// Mitsubishi GX Works2 project: B_v6_v2   PLC: Q03UDE

PROGRAM COMMON
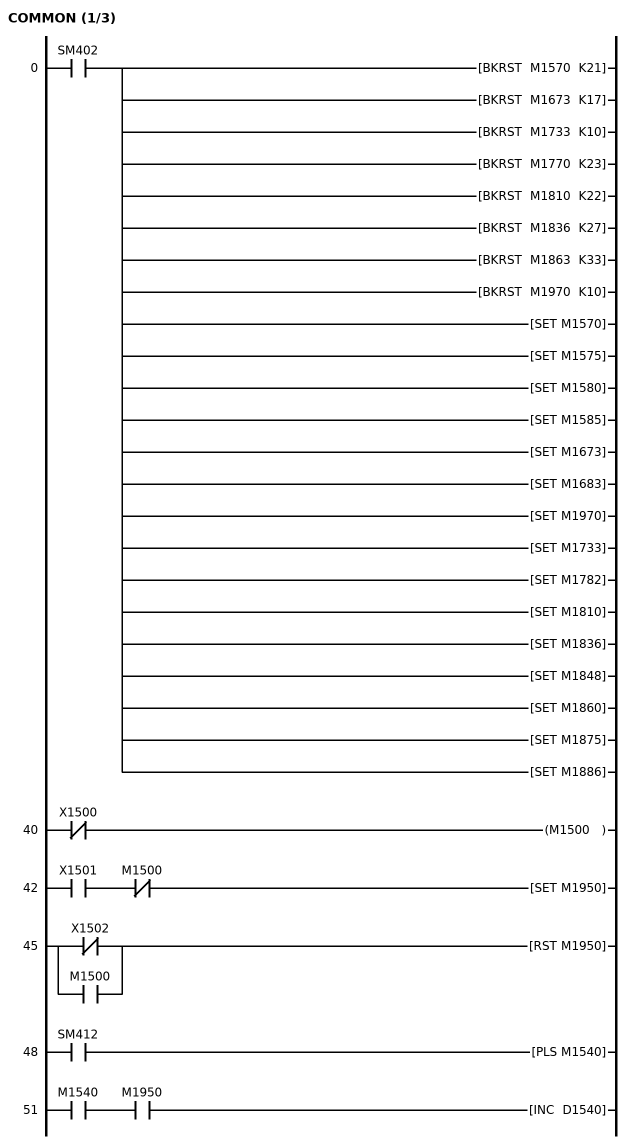
0     LD      SM402
      BKRST   M1570 K21
      BKRST   M1673 K17
      BKRST   M1733 K10
      BKRST   M1770 K23
      BKRST   M1810 K22
      BKRST   M1836 K27
      BKRST   M1863 K33
      BKRST   M1970 K10
      SET     M1570
      SET     M1575
      SET     M1580
      SET     M1585
      SET     M1673
      SET     M1683
      SET     M1970
      SET     M1733
      SET     M1782
      SET     M1810
      SET     M1836
      SET     M1848
      SET     M1860
      SET     M1875
      SET     M1886
40    LDI     X1500
      OUT     M1500
42    LD      X1501
      ANI     M1500
      SET     M1950
45    LDI     X1502
      OR      M1500
      RST     M1950
48    LD      SM412
      PLS     M1540
51    LD      M1540
      AND     M1950
      INC     D1540
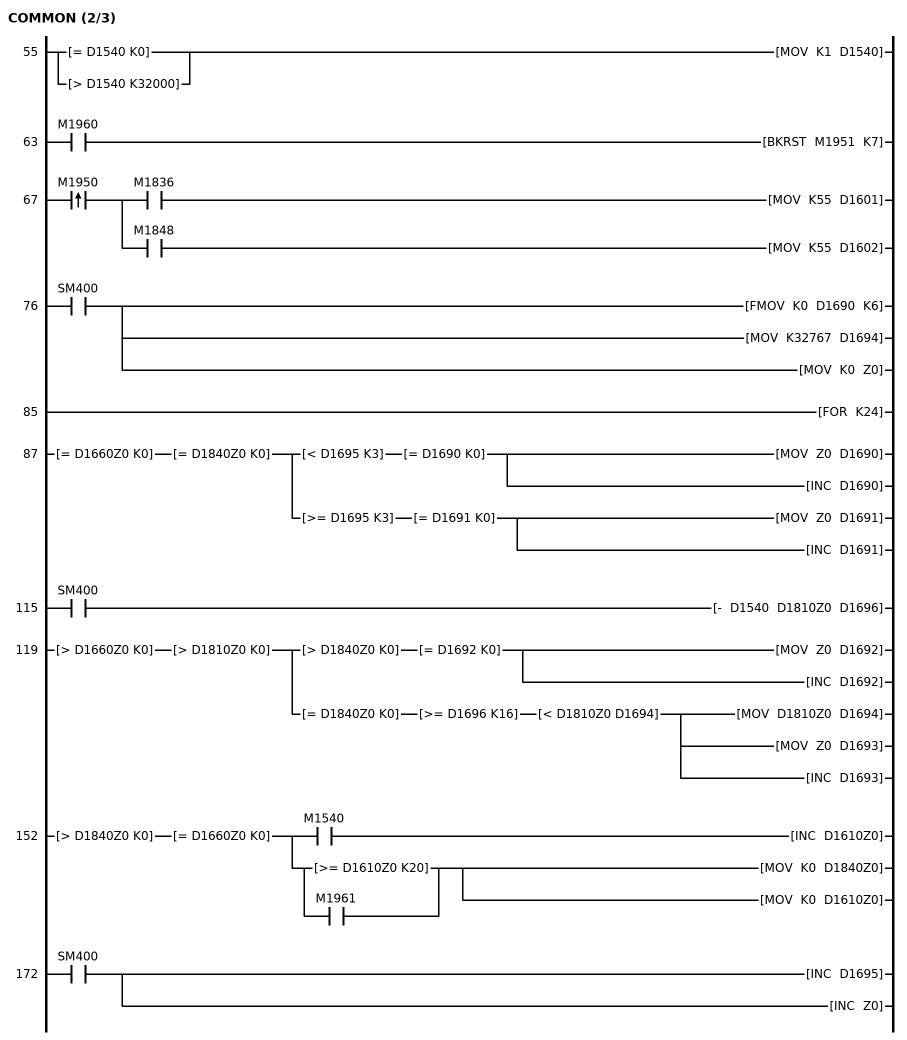
55    LD=     D1540 K0
      OR>     D1540 K32000
      MOV     K1 D1540
63    LD      M1960
      BKRST   M1951 K7
67    LDP     M1950
      MPS
      AND     M1836
      MOV     K55 D1601
      MPP
      AND     M1848
      MOV     K55 D1602
76    LD      SM400
      FMOV    K0 D1690 K6
      MOV     K32767 D1694
      MOV     K0 Z0
85    FOR     K24
87    LD=     D1660Z0 K0
      AND=    D1840Z0 K0
      MPS
      AND<    D1695 K3
      AND=    D1690 K0
      MOV     Z0 D1690
      INC     D1690
      MPP
      AND>=   D1695 K3
      AND=    D1691 K0
      MOV     Z0 D1691
      INC     D1691
115   LD      SM400
      -       D1540 D1810Z0 D1696
119   LD>     D1660Z0 K0
      AND>    D1810Z0 K0
      MPS
      AND>    D1840Z0 K0
      AND=    D1692 K0
      MOV     Z0 D1692
      INC     D1692
      MPP
      AND=    D1840Z0 K0
      AND>=   D1696 K16
      AND<    D1810Z0 D1694
      MOV     D1810Z0 D1694
      MOV     Z0 D1693
      INC     D1693
152   LD>     D1840Z0 K0
      AND=    D1660Z0 K0
      MPS
      AND     M1540
      INC     D1610Z0
      MPP
      LD>=    D1610Z0 K20
      OR      M1961
      ANB
      MOV     K0 D1840Z0
      MOV     K0 D1610Z0
172   LD      SM400
      INC     D1695
      INC     Z0
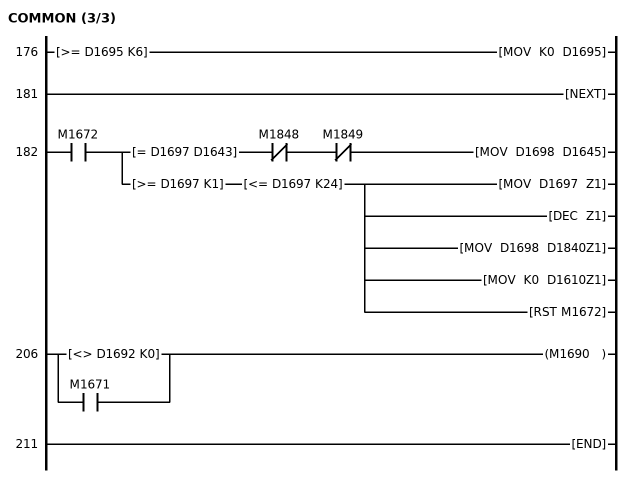
176   LD>=    D1695 K6
      MOV     K0 D1695
181   NEXT
182   LD      M1672
      MPS
      AND=    D1697 D1643
      ANI     M1848
      ANI     M1849
      MOV     D1698 D1645
      MPP
      AND>=   D1697 K1
      AND<=   D1697 K24
      MOV     D1697 Z1
      DEC     Z1
      MOV     D1698 D1840Z1
      MOV     K0 D1610Z1
      RST     M1672
206   LD<>    D1692 K0
      OR      M1671
      OUT     M1690
211   END
END_PROGRAM

PROGRAM RFID
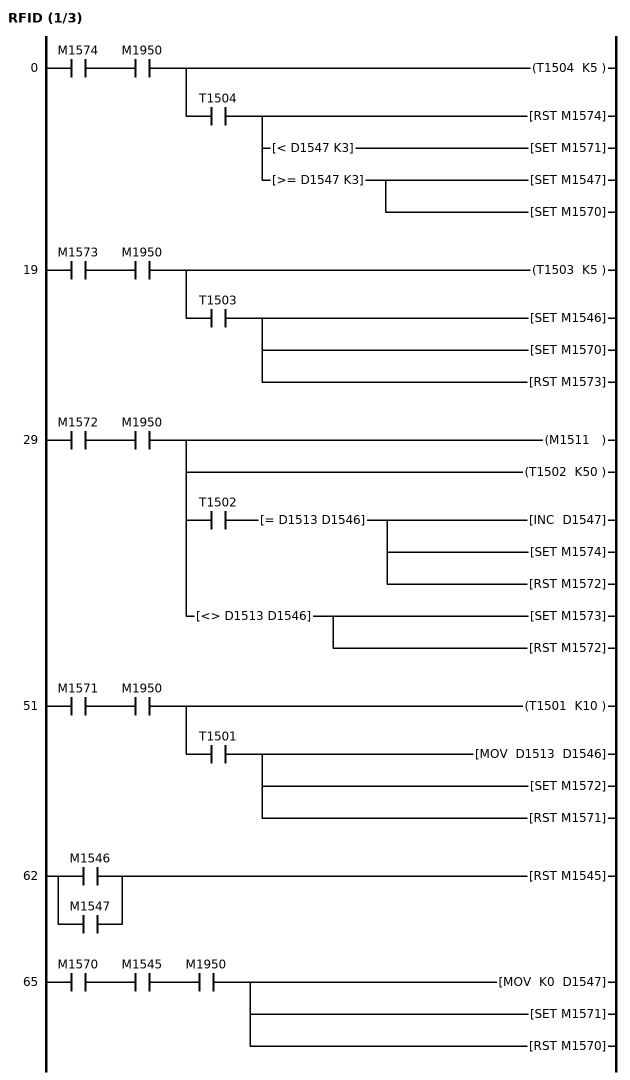
0     LD      M1574
      AND     M1950
      OUT     T1504 K5
      AND     T1504
      RST     M1574
      MPS
      AND<    D1547 K3
      SET     M1571
      MPP
      AND>=   D1547 K3
      SET     M1547
      SET     M1570
19    LD      M1573
      AND     M1950
      OUT     T1503 K5
      AND     T1503
      SET     M1546
      SET     M1570
      RST     M1573
29    LD      M1572
      AND     M1950
      OUT     M1511
      OUT     T1502 K50
      MPS
      AND     T1502
      AND=    D1513 D1546
      INC     D1547
      SET     M1574
      RST     M1572
      MPP
      AND<>   D1513 D1546
      SET     M1573
      RST     M1572
51    LD      M1571
      AND     M1950
      OUT     T1501 K10
      AND     T1501
      MOV     D1513 D1546
      SET     M1572
      RST     M1571
62    LD      M1546
      OR      M1547
      RST     M1545
65    LD      M1570
      AND     M1545
      AND     M1950
      MOV     K0 D1547
      SET     M1571
      RST     M1570
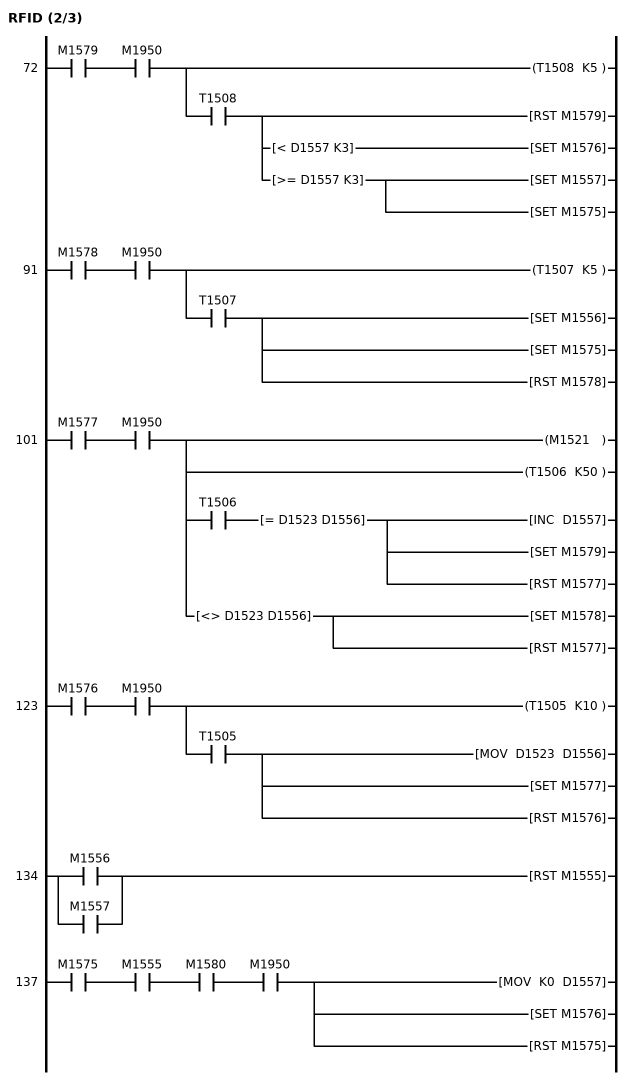
72    LD      M1579
      AND     M1950
      OUT     T1508 K5
      AND     T1508
      RST     M1579
      MPS
      AND<    D1557 K3
      SET     M1576
      MPP
      AND>=   D1557 K3
      SET     M1557
      SET     M1575
91    LD      M1578
      AND     M1950
      OUT     T1507 K5
      AND     T1507
      SET     M1556
      SET     M1575
      RST     M1578
101   LD      M1577
      AND     M1950
      OUT     M1521
      OUT     T1506 K50
      MPS
      AND     T1506
      AND=    D1523 D1556
      INC     D1557
      SET     M1579
      RST     M1577
      MPP
      AND<>   D1523 D1556
      SET     M1578
      RST     M1577
123   LD      M1576
      AND     M1950
      OUT     T1505 K10
      AND     T1505
      MOV     D1523 D1556
      SET     M1577
      RST     M1576
134   LD      M1556
      OR      M1557
      RST     M1555
137   LD      M1575
      AND     M1555
      AND     M1580
      AND     M1950
      MOV     K0 D1557
      SET     M1576
      RST     M1575
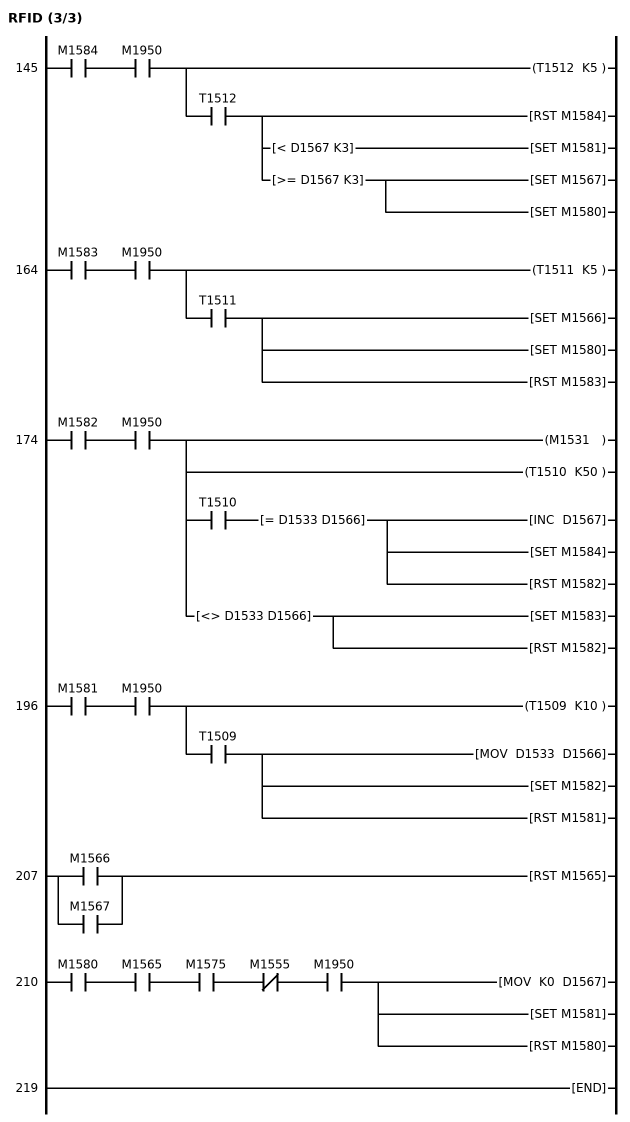
145   LD      M1584
      AND     M1950
      OUT     T1512 K5
      AND     T1512
      RST     M1584
      MPS
      AND<    D1567 K3
      SET     M1581
      MPP
      AND>=   D1567 K3
      SET     M1567
      SET     M1580
164   LD      M1583
      AND     M1950
      OUT     T1511 K5
      AND     T1511
      SET     M1566
      SET     M1580
      RST     M1583
174   LD      M1582
      AND     M1950
      OUT     M1531
      OUT     T1510 K50
      MPS
      AND     T1510
      AND=    D1533 D1566
      INC     D1567
      SET     M1584
      RST     M1582
      MPP
      AND<>   D1533 D1566
      SET     M1583
      RST     M1582
196   LD      M1581
      AND     M1950
      OUT     T1509 K10
      AND     T1509
      MOV     D1533 D1566
      SET     M1582
      RST     M1581
207   LD      M1566
      OR      M1567
      RST     M1565
210   LD      M1580
      AND     M1565
      AND     M1575
      ANI     M1555
      AND     M1950
      MOV     K0 D1567
      SET     M1581
      RST     M1580
219   END
END_PROGRAM

PROGRAM INFEED
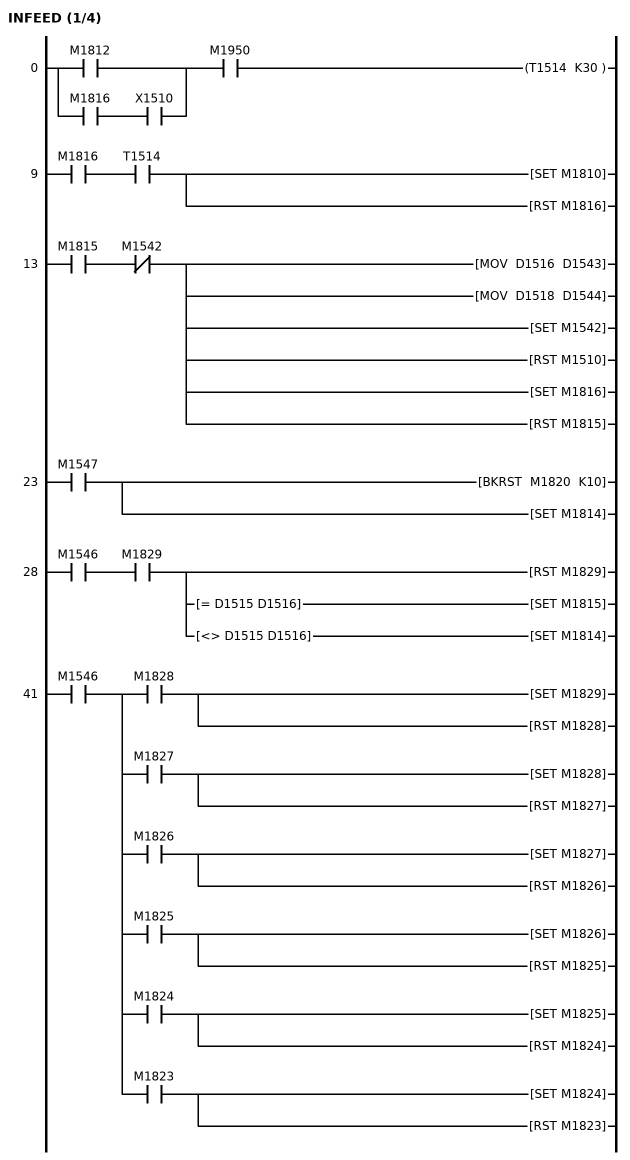
0     LD      M1812
      LD      M1816
      AND     X1510
      ORB
      AND     M1950
      OUT     T1514 K30
9     LD      M1816
      AND     T1514
      SET     M1810
      RST     M1816
13    LD      M1815
      ANI     M1542
      MOV     D1516 D1543
      MOV     D1518 D1544
      SET     M1542
      RST     M1510
      SET     M1816
      RST     M1815
23    LD      M1547
      BKRST   M1820 K10
      SET     M1814
28    LD      M1546
      AND     M1829
      RST     M1829
      MPS
      AND=    D1515 D1516
      SET     M1815
      MPP
      AND<>   D1515 D1516
      SET     M1814
41    LD      M1546
      MPS
      AND     M1828
      SET     M1829
      RST     M1828
      MRD
      AND     M1827
      SET     M1828
      RST     M1827
      MRD
      AND     M1826
      SET     M1827
      RST     M1826
      MRD
      AND     M1825
      SET     M1826
      RST     M1825
      MRD
      AND     M1824
      SET     M1825
      RST     M1824
      MPP
      AND     M1823
      SET     M1824
      RST     M1823
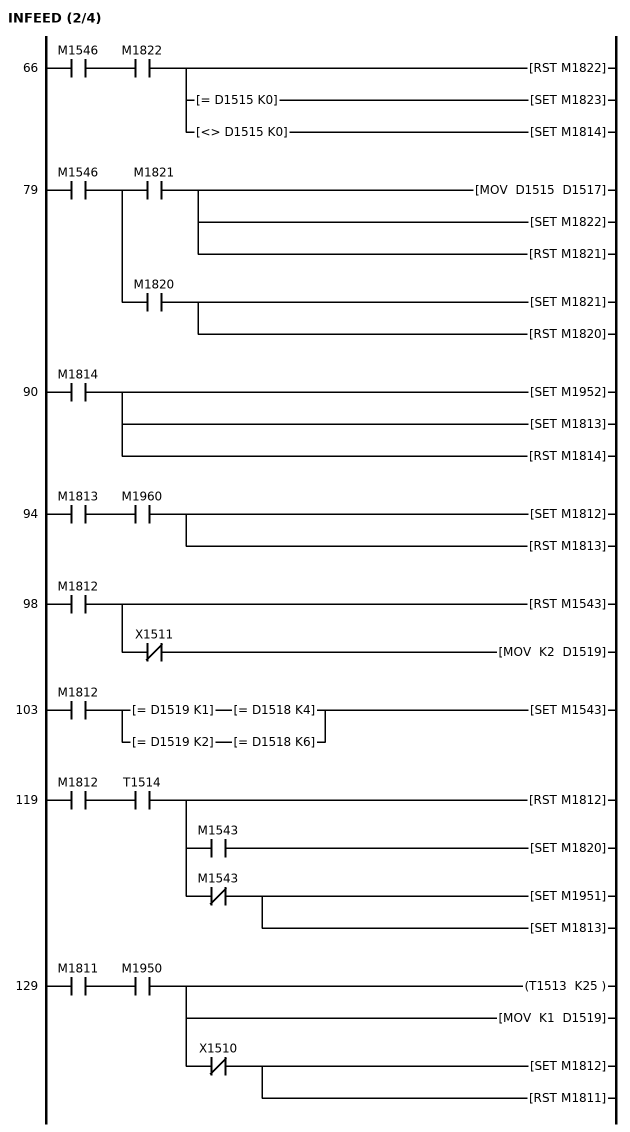
66    LD      M1546
      AND     M1822
      RST     M1822
      MPS
      AND=    D1515 K0
      SET     M1823
      MPP
      AND<>   D1515 K0
      SET     M1814
79    LD      M1546
      MPS
      AND     M1821
      MOV     D1515 D1517
      SET     M1822
      RST     M1821
      MPP
      AND     M1820
      SET     M1821
      RST     M1820
90    LD      M1814
      SET     M1952
      SET     M1813
      RST     M1814
94    LD      M1813
      AND     M1960
      SET     M1812
      RST     M1813
98    LD      M1812
      RST     M1543
      ANI     X1511
      MOV     K2 D1519
103   LD      M1812
      LD=     D1519 K1
      AND=    D1518 K4
      LD=     D1519 K2
      AND=    D1518 K6
      ORB
      ANB
      SET     M1543
119   LD      M1812
      AND     T1514
      RST     M1812
      MPS
      AND     M1543
      SET     M1820
      MPP
      ANI     M1543
      SET     M1951
      SET     M1813
129   LD      M1811
      AND     M1950
      OUT     T1513 K25
      MOV     K1 D1519
      ANI     X1510
      SET     M1812
      RST     M1811
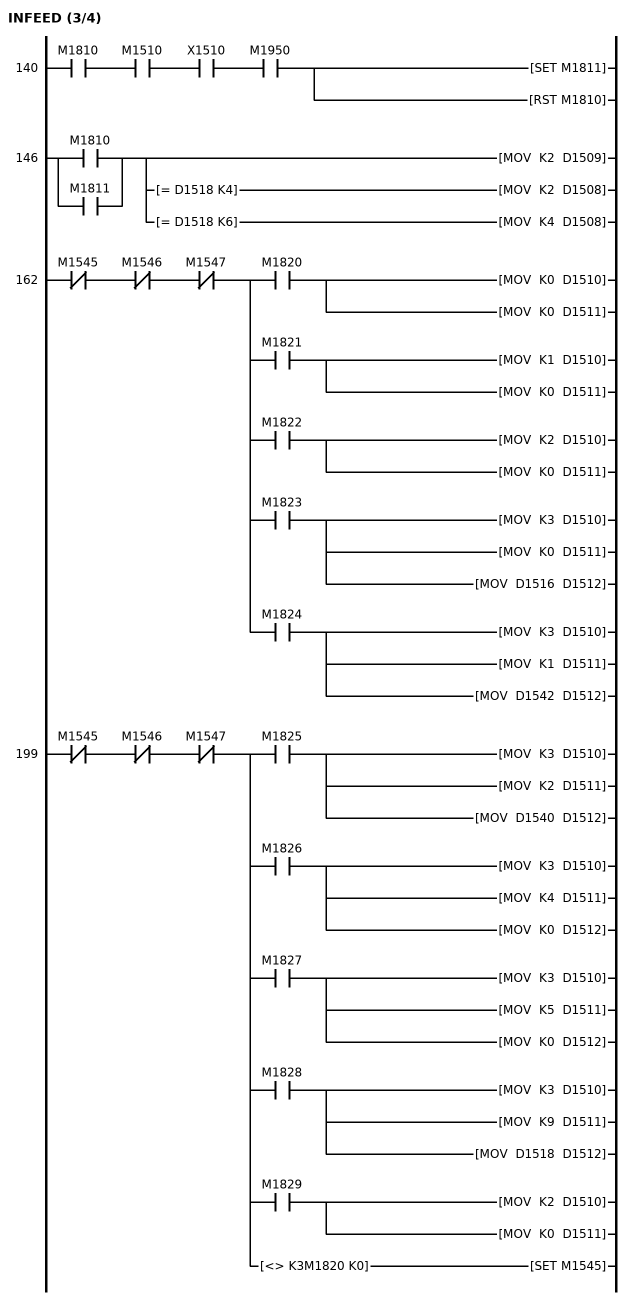
140   LD      M1810
      AND     M1510
      AND     X1510
      AND     M1950
      SET     M1811
      RST     M1810
146   LD      M1810
      OR      M1811
      MOV     K2 D1509
      MPS
      AND=    D1518 K4
      MOV     K2 D1508
      MPP
      AND=    D1518 K6
      MOV     K4 D1508
162   LDI     M1545
      ANI     M1546
      ANI     M1547
      MPS
      AND     M1820
      MOV     K0 D1510
      MOV     K0 D1511
      MRD
      AND     M1821
      MOV     K1 D1510
      MOV     K0 D1511
      MRD
      AND     M1822
      MOV     K2 D1510
      MOV     K0 D1511
      MRD
      AND     M1823
      MOV     K3 D1510
      MOV     K0 D1511
      MOV     D1516 D1512
      MPP
      AND     M1824
      MOV     K3 D1510
      MOV     K1 D1511
      MOV     D1542 D1512
199   LDI     M1545
      ANI     M1546
      ANI     M1547
      MPS
      AND     M1825
      MOV     K3 D1510
      MOV     K2 D1511
      MOV     D1540 D1512
      MRD
      AND     M1826
      MOV     K3 D1510
      MOV     K4 D1511
      MOV     K0 D1512
      MRD
      AND     M1827
      MOV     K3 D1510
      MOV     K5 D1511
      MOV     K0 D1512
      MRD
      AND     M1828
      MOV     K3 D1510
      MOV     K9 D1511
      MOV     D1518 D1512
      MRD
      AND     M1829
      MOV     K2 D1510
      MOV     K0 D1511
      MPP
      AND<>   K3M1820 K0
      SET     M1545
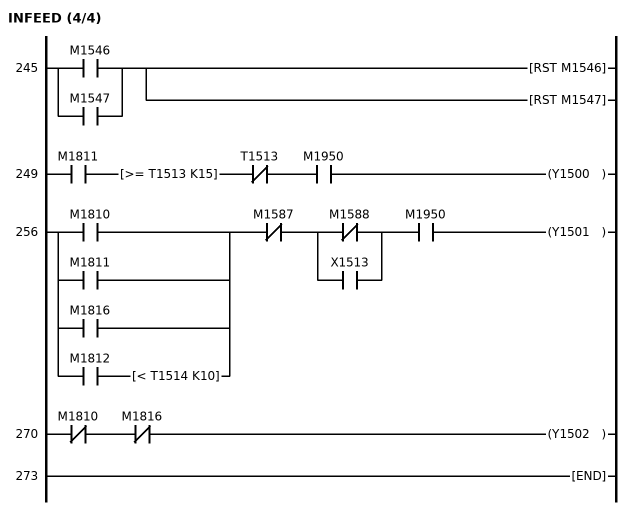
245   LD      M1546
      OR      M1547
      RST     M1546
      RST     M1547
249   LD      M1811
      AND>=   T1513 K15
      ANI     T1513
      AND     M1950
      OUT     Y1500
256   LD      M1810
      OR      M1811
      OR      M1816
      LD      M1812
      AND<    T1514 K10
      ORB
      ANI     M1587
      LDI     M1588
      OR      X1513
      ANB
      AND     M1950
      OUT     Y1501
270   LDI     M1810
      ANI     M1816
      OUT     Y1502
273   END
END_PROGRAM

PROGRAM CRANE
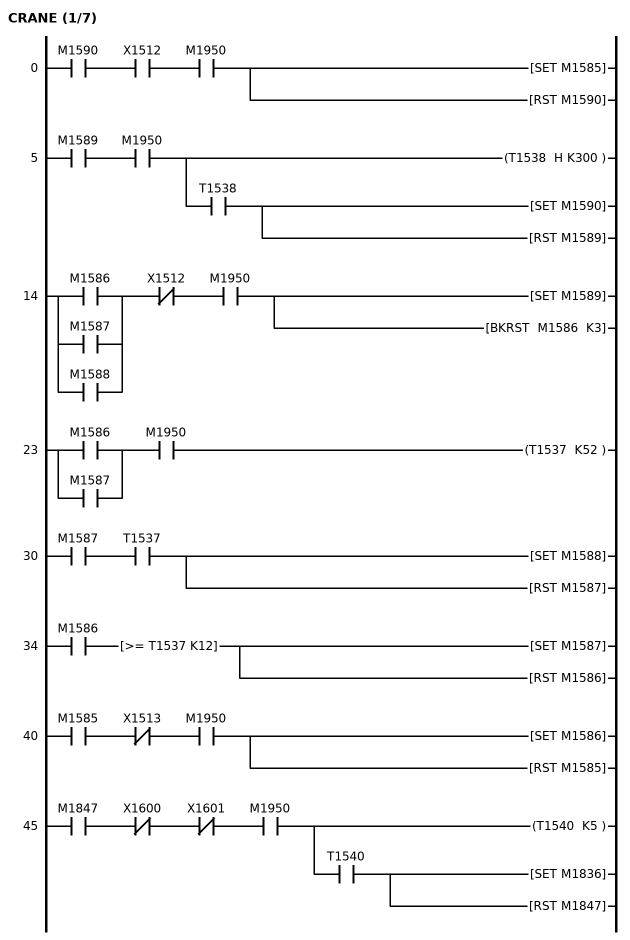
0     LD      M1590
      AND     X1512
      AND     M1950
      SET     M1585
      RST     M1590
5     LD      M1589
      AND     M1950
      OUTH    T1538 K300
      AND     T1538
      SET     M1590
      RST     M1589
14    LD      M1586
      OR      M1587
      OR      M1588
      ANI     X1512
      AND     M1950
      SET     M1589
      BKRST   M1586 K3
23    LD      M1586
      OR      M1587
      AND     M1950
      OUT     T1537 K52
30    LD      M1587
      AND     T1537
      SET     M1588
      RST     M1587
34    LD      M1586
      AND>=   T1537 K12
      SET     M1587
      RST     M1586
40    LD      M1585
      ANI     X1513
      AND     M1950
      SET     M1586
      RST     M1585
45    LD      M1847
      ANI     X1600
      ANI     X1601
      AND     M1950
      OUT     T1540 K5
      AND     T1540
      SET     M1836
      RST     M1847
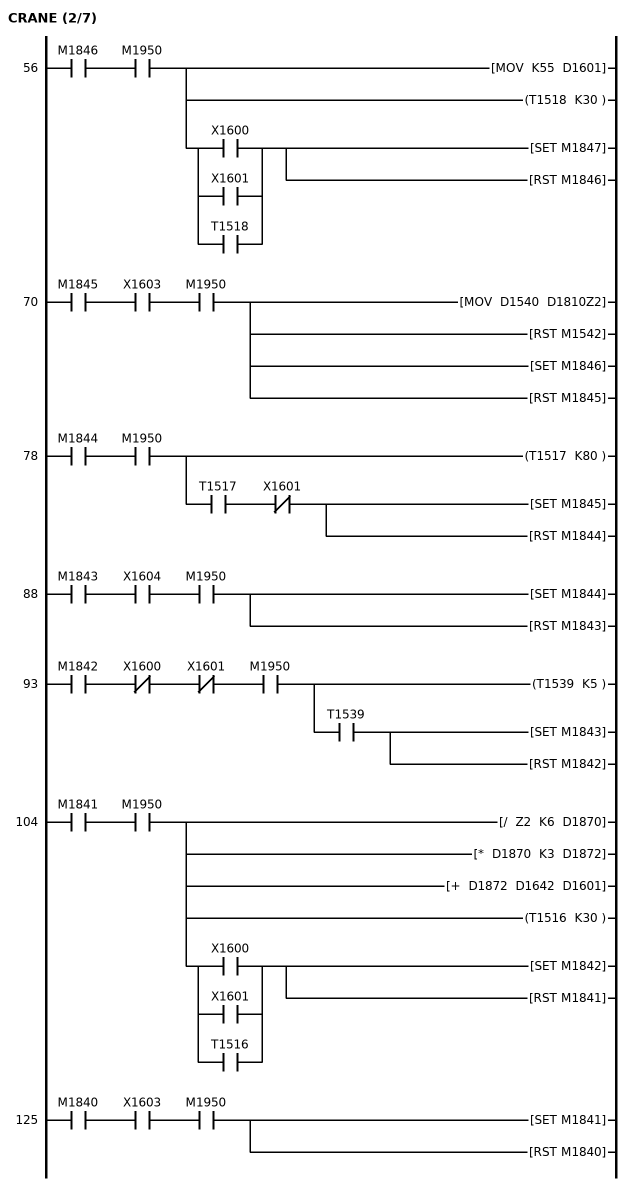
56    LD      M1846
      AND     M1950
      MOV     K55 D1601
      OUT     T1518 K30
      LD      X1600
      OR      X1601
      OR      T1518
      ANB
      SET     M1847
      RST     M1846
70    LD      M1845
      AND     X1603
      AND     M1950
      MOV     D1540 D1810Z2
      RST     M1542
      SET     M1846
      RST     M1845
78    LD      M1844
      AND     M1950
      OUT     T1517 K80
      AND     T1517
      ANI     X1601
      SET     M1845
      RST     M1844
88    LD      M1843
      AND     X1604
      AND     M1950
      SET     M1844
      RST     M1843
93    LD      M1842
      ANI     X1600
      ANI     X1601
      AND     M1950
      OUT     T1539 K5
      AND     T1539
      SET     M1843
      RST     M1842
104   LD      M1841
      AND     M1950
      /       Z2 K6 D1870
      *       D1870 K3 D1872
      +       D1872 D1642 D1601
      OUT     T1516 K30
      LD      X1600
      OR      X1601
      OR      T1516
      ANB
      SET     M1842
      RST     M1841
125   LD      M1840
      AND     X1603
      AND     M1950
      SET     M1841
      RST     M1840
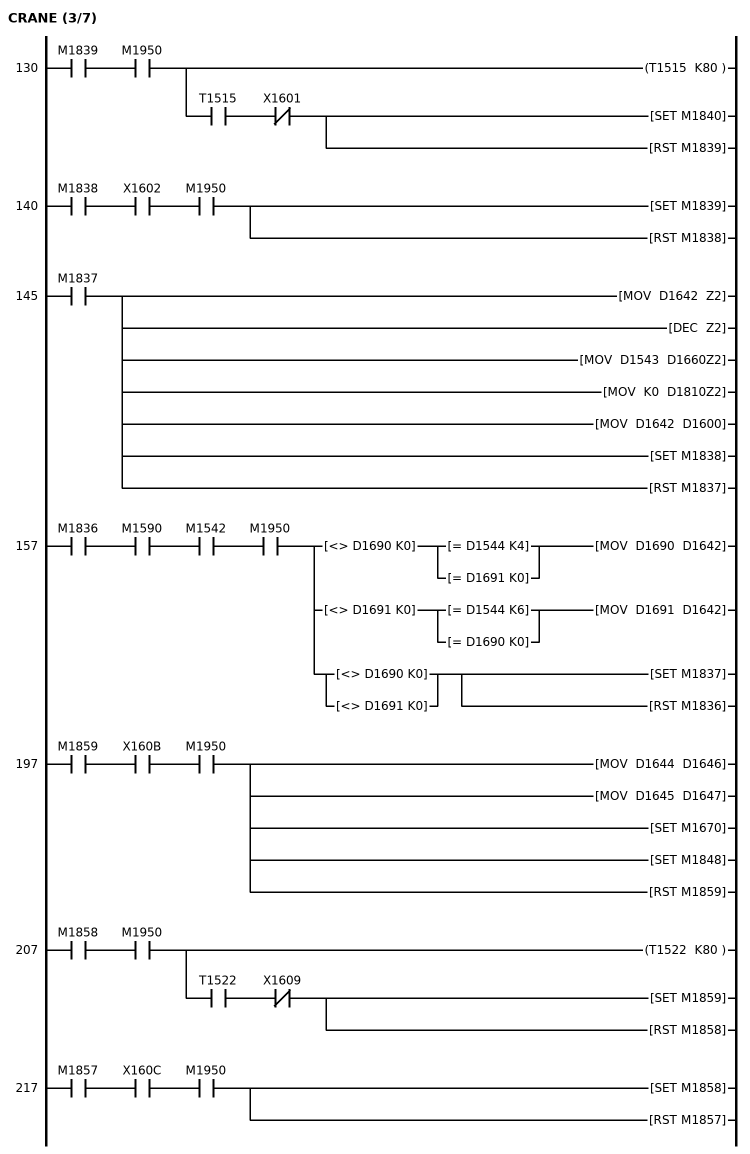
130   LD      M1839
      AND     M1950
      OUT     T1515 K80
      AND     T1515
      ANI     X1601
      SET     M1840
      RST     M1839
140   LD      M1838
      AND     X1602
      AND     M1950
      SET     M1839
      RST     M1838
145   LD      M1837
      MOV     D1642 Z2
      DEC     Z2
      MOV     D1543 D1660Z2
      MOV     K0 D1810Z2
      MOV     D1642 D1600
      SET     M1838
      RST     M1837
157   LD      M1836
      AND     M1590
      AND     M1542
      AND     M1950
      MPS
      AND<>   D1690 K0
      LD=     D1544 K4
      OR=     D1691 K0
      ANB
      MOV     D1690 D1642
      MRD
      AND<>   D1691 K0
      LD=     D1544 K6
      OR=     D1690 K0
      ANB
      MOV     D1691 D1642
      MPP
      LD<>    D1690 K0
      OR<>    D1691 K0
      ANB
      SET     M1837
      RST     M1836
197   LD      M1859
      AND     X160B
      AND     M1950
      MOV     D1644 D1646
      MOV     D1645 D1647
      SET     M1670
      SET     M1848
      RST     M1859
207   LD      M1858
      AND     M1950
      OUT     T1522 K80
      AND     T1522
      ANI     X1609
      SET     M1859
      RST     M1858
217   LD      M1857
      AND     X160C
      AND     M1950
      SET     M1858
      RST     M1857
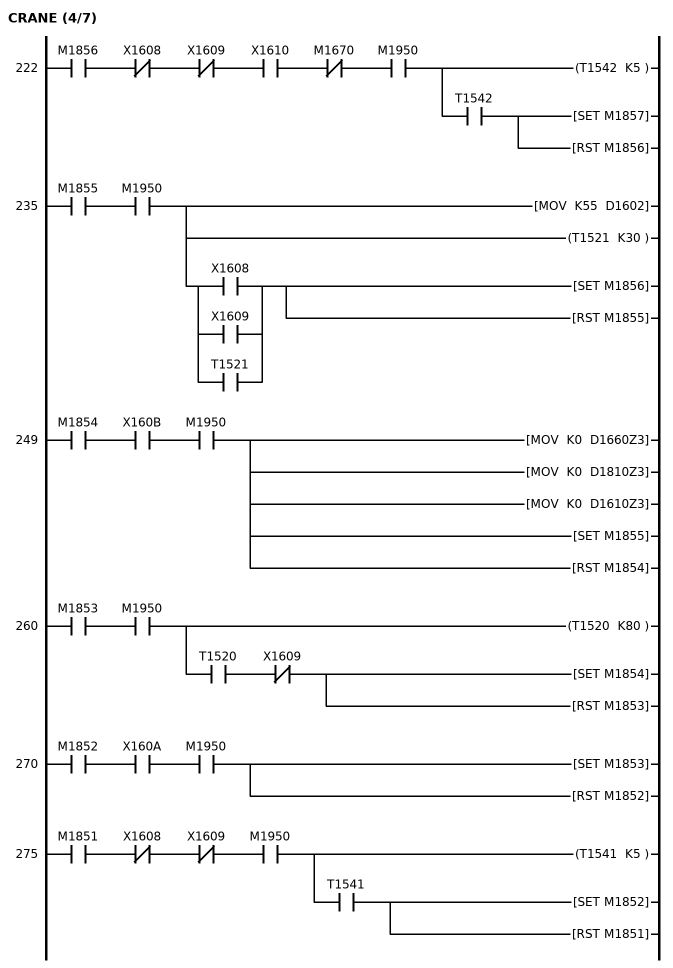
222   LD      M1856
      ANI     X1608
      ANI     X1609
      AND     X1610
      ANI     M1670
      AND     M1950
      OUT     T1542 K5
      AND     T1542
      SET     M1857
      RST     M1856
235   LD      M1855
      AND     M1950
      MOV     K55 D1602
      OUT     T1521 K30
      LD      X1608
      OR      X1609
      OR      T1521
      ANB
      SET     M1856
      RST     M1855
249   LD      M1854
      AND     X160B
      AND     M1950
      MOV     K0 D1660Z3
      MOV     K0 D1810Z3
      MOV     K0 D1610Z3
      SET     M1855
      RST     M1854
260   LD      M1853
      AND     M1950
      OUT     T1520 K80
      AND     T1520
      ANI     X1609
      SET     M1854
      RST     M1853
270   LD      M1852
      AND     X160A
      AND     M1950
      SET     M1853
      RST     M1852
275   LD      M1851
      ANI     X1608
      ANI     X1609
      AND     M1950
      OUT     T1541 K5
      AND     T1541
      SET     M1852
      RST     M1851
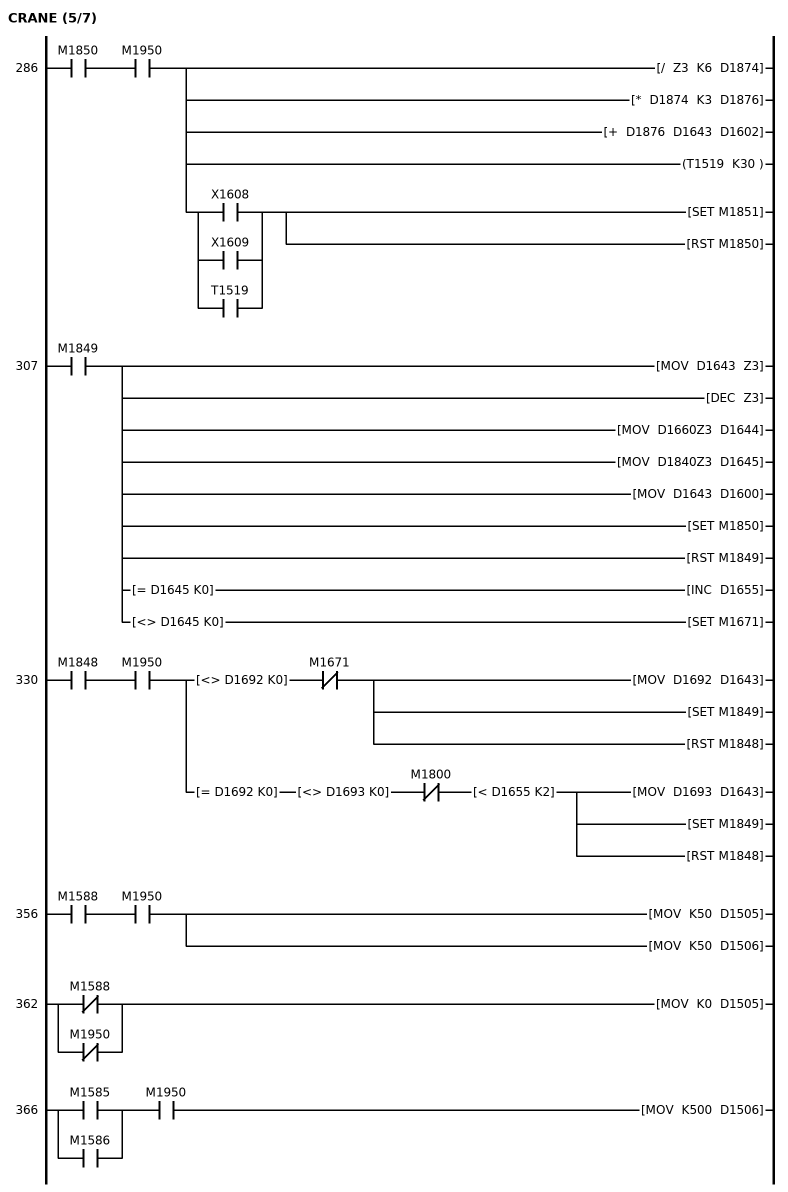
286   LD      M1850
      AND     M1950
      /       Z3 K6 D1874
      *       D1874 K3 D1876
      +       D1876 D1643 D1602
      OUT     T1519 K30
      LD      X1608
      OR      X1609
      OR      T1519
      ANB
      SET     M1851
      RST     M1850
307   LD      M1849
      MOV     D1643 Z3
      DEC     Z3
      MOV     D1660Z3 D1644
      MOV     D1840Z3 D1645
      MOV     D1643 D1600
      SET     M1850
      RST     M1849
      MPS
      AND=    D1645 K0
      INC     D1655
      MPP
      AND<>   D1645 K0
      SET     M1671
330   LD      M1848
      AND     M1950
      MPS
      AND<>   D1692 K0
      ANI     M1671
      MOV     D1692 D1643
      SET     M1849
      RST     M1848
      MPP
      AND=    D1692 K0
      AND<>   D1693 K0
      ANI     M1800
      AND<    D1655 K2
      MOV     D1693 D1643
      SET     M1849
      RST     M1848
356   LD      M1588
      AND     M1950
      MOV     K50 D1505
      MOV     K50 D1506
362   LDI     M1588
      ORI     M1950
      MOV     K0 D1505
366   LD      M1585
      OR      M1586
      AND     M1950
      MOV     K500 D1506
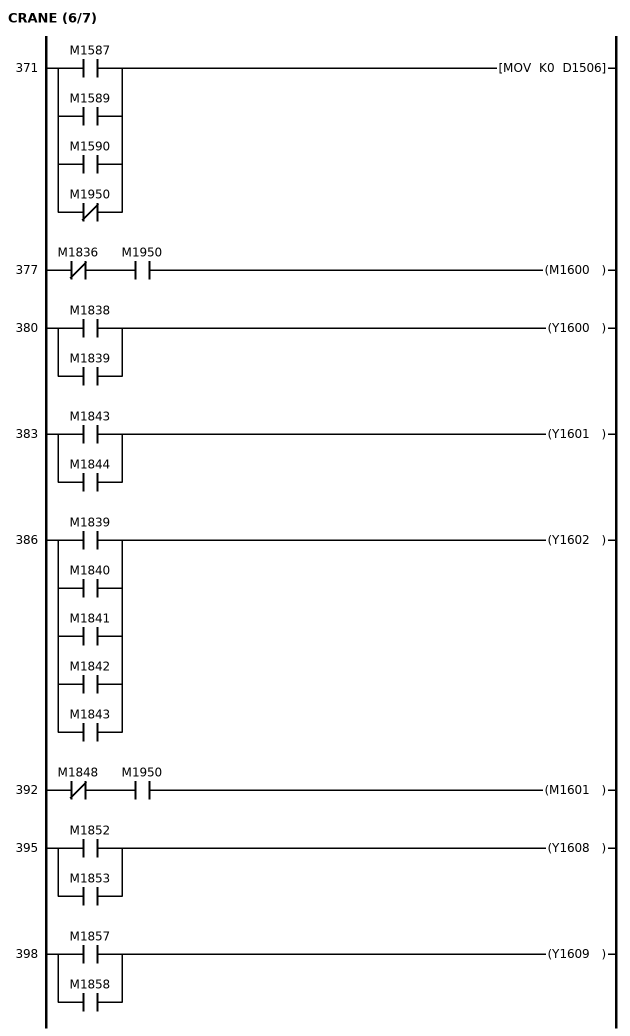
371   LD      M1587
      OR      M1589
      OR      M1590
      ORI     M1950
      MOV     K0 D1506
377   LDI     M1836
      AND     M1950
      OUT     M1600
380   LD      M1838
      OR      M1839
      OUT     Y1600
383   LD      M1843
      OR      M1844
      OUT     Y1601
386   LD      M1839
      OR      M1840
      OR      M1841
      OR      M1842
      OR      M1843
      OUT     Y1602
392   LDI     M1848
      AND     M1950
      OUT     M1601
395   LD      M1852
      OR      M1853
      OUT     Y1608
398   LD      M1857
      OR      M1858
      OUT     Y1609
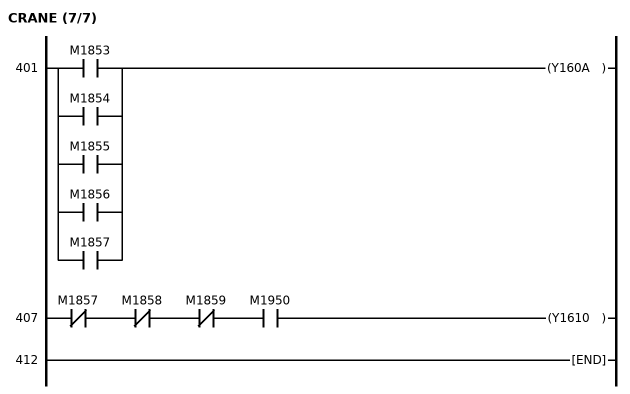
401   LD      M1853
      OR      M1854
      OR      M1855
      OR      M1856
      OR      M1857
      OUT     Y160A
407   LDI     M1857
      ANI     M1858
      ANI     M1859
      AND     M1950
      OUT     Y1610
412   END
END_PROGRAM

PROGRAM SORT1
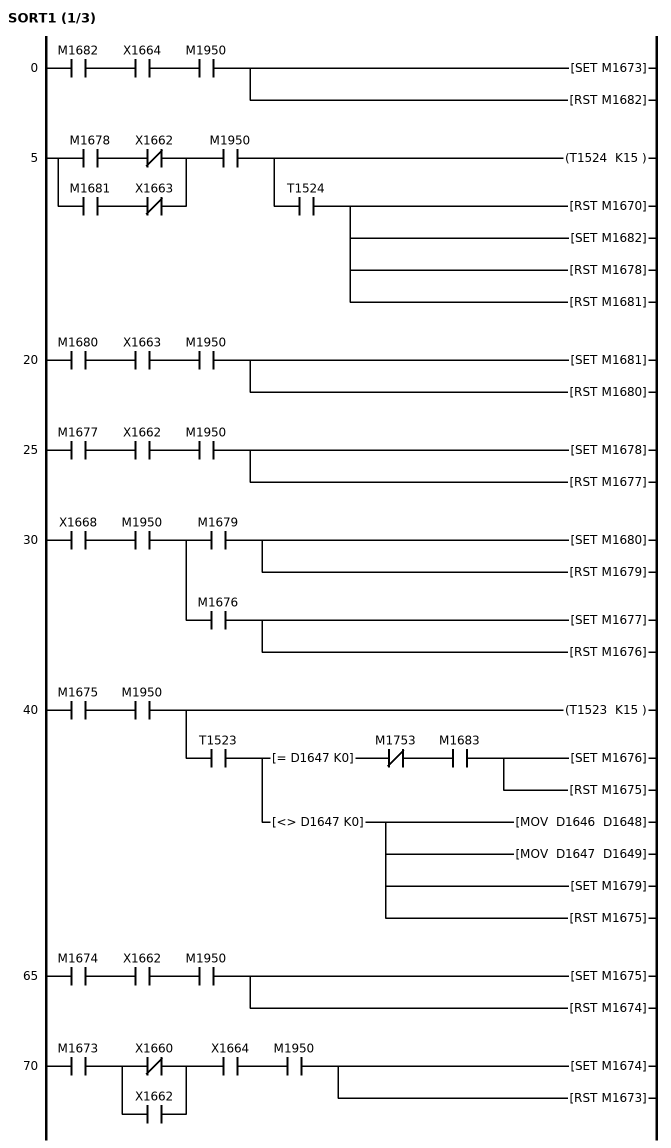
0     LD      M1682
      AND     X1664
      AND     M1950
      SET     M1673
      RST     M1682
5     LD      M1678
      ANI     X1662
      LD      M1681
      ANI     X1663
      ORB
      AND     M1950
      OUT     T1524 K15
      AND     T1524
      RST     M1670
      SET     M1682
      RST     M1678
      RST     M1681
20    LD      M1680
      AND     X1663
      AND     M1950
      SET     M1681
      RST     M1680
25    LD      M1677
      AND     X1662
      AND     M1950
      SET     M1678
      RST     M1677
30    LD      X1668
      AND     M1950
      MPS
      AND     M1679
      SET     M1680
      RST     M1679
      MPP
      AND     M1676
      SET     M1677
      RST     M1676
40    LD      M1675
      AND     M1950
      OUT     T1523 K15
      AND     T1523
      MPS
      AND=    D1647 K0
      ANI     M1753
      AND     M1683
      SET     M1676
      RST     M1675
      MPP
      AND<>   D1647 K0
      MOV     D1646 D1648
      MOV     D1647 D1649
      SET     M1679
      RST     M1675
65    LD      M1674
      AND     X1662
      AND     M1950
      SET     M1675
      RST     M1674
70    LD      M1673
      LDI     X1660
      OR      X1662
      ANB
      AND     X1664
      AND     M1950
      SET     M1674
      RST     M1673
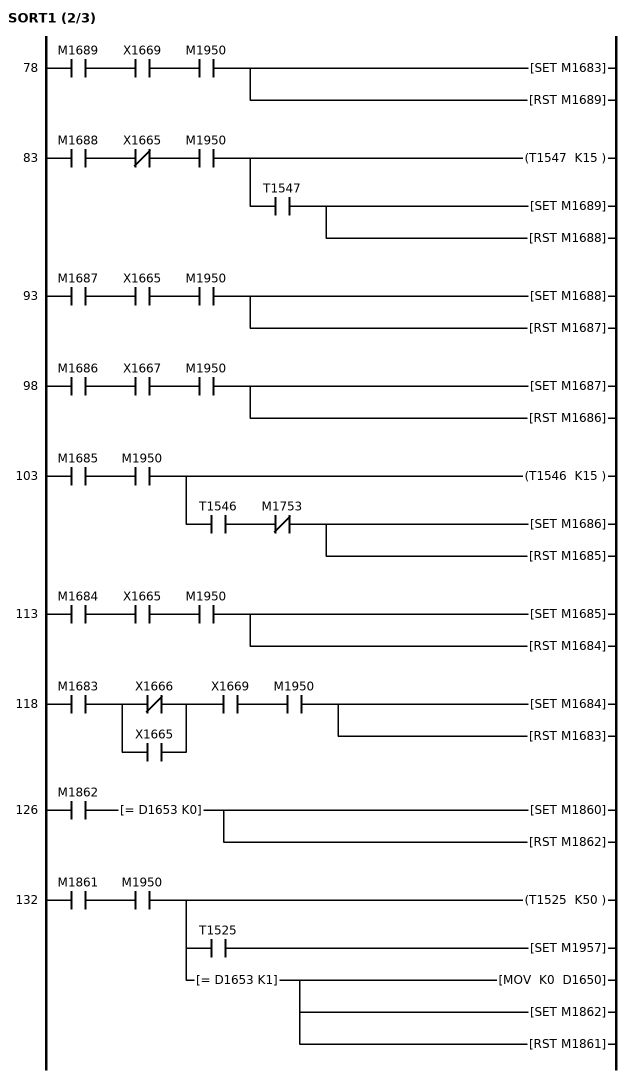
78    LD      M1689
      AND     X1669
      AND     M1950
      SET     M1683
      RST     M1689
83    LD      M1688
      ANI     X1665
      AND     M1950
      OUT     T1547 K15
      AND     T1547
      SET     M1689
      RST     M1688
93    LD      M1687
      AND     X1665
      AND     M1950
      SET     M1688
      RST     M1687
98    LD      M1686
      AND     X1667
      AND     M1950
      SET     M1687
      RST     M1686
103   LD      M1685
      AND     M1950
      OUT     T1546 K15
      AND     T1546
      ANI     M1753
      SET     M1686
      RST     M1685
113   LD      M1684
      AND     X1665
      AND     M1950
      SET     M1685
      RST     M1684
118   LD      M1683
      LDI     X1666
      OR      X1665
      ANB
      AND     X1669
      AND     M1950
      SET     M1684
      RST     M1683
126   LD      M1862
      AND=    D1653 K0
      SET     M1860
      RST     M1862
132   LD      M1861
      AND     M1950
      OUT     T1525 K50
      MPS
      AND     T1525
      SET     M1957
      MPP
      AND=    D1653 K1
      MOV     K0 D1650
      SET     M1862
      RST     M1861
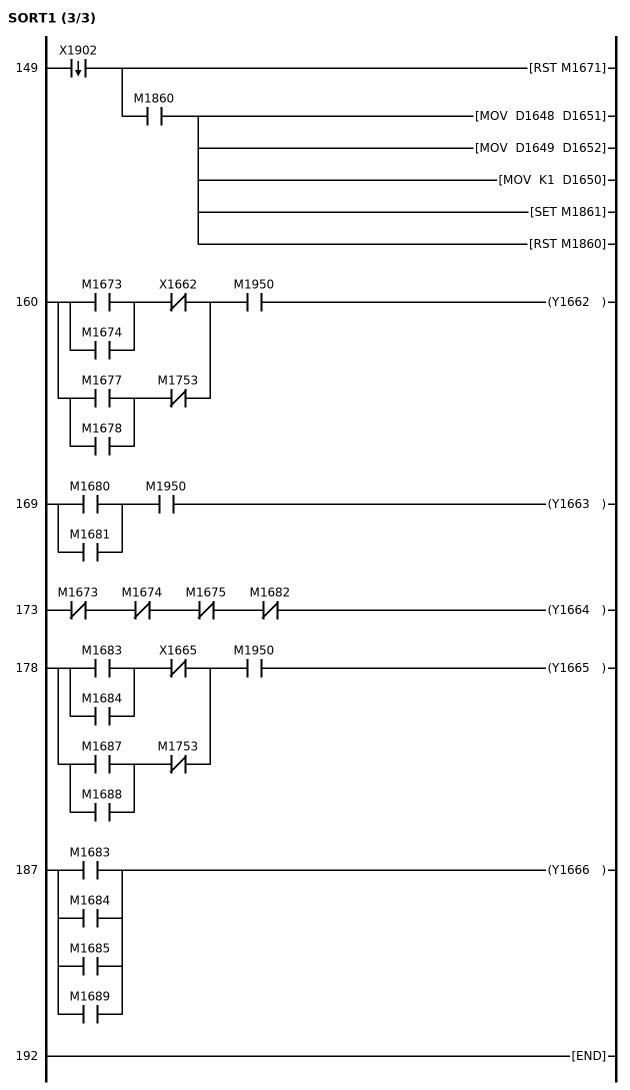
149   LDF     X1902
      RST     M1671
      AND     M1860
      MOV     D1648 D1651
      MOV     D1649 D1652
      MOV     K1 D1650
      SET     M1861
      RST     M1860
160   LD      M1673
      OR      M1674
      ANI     X1662
      LD      M1677
      OR      M1678
      ANI     M1753
      ORB
      AND     M1950
      OUT     Y1662
169   LD      M1680
      OR      M1681
      AND     M1950
      OUT     Y1663
173   LDI     M1673
      ANI     M1674
      ANI     M1675
      ANI     M1682
      OUT     Y1664
178   LD      M1683
      OR      M1684
      ANI     X1665
      LD      M1687
      OR      M1688
      ANI     M1753
      ORB
      AND     M1950
      OUT     Y1665
187   LD      M1683
      OR      M1684
      OR      M1685
      OR      M1689
      OUT     Y1666
192   END
END_PROGRAM

PROGRAM INSPECT
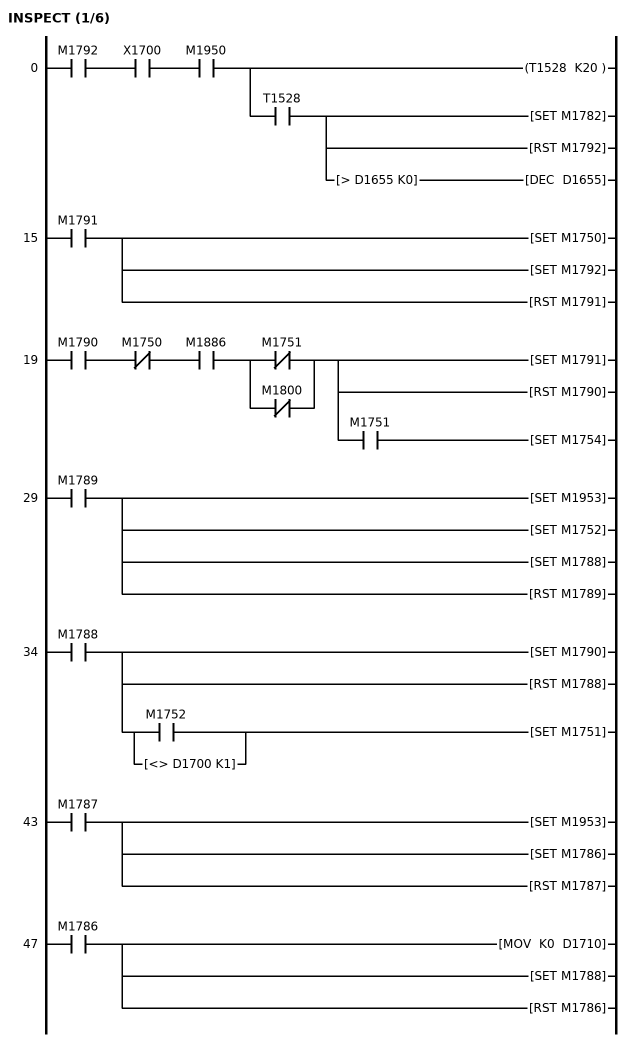
0     LD      M1792
      AND     X1700
      AND     M1950
      OUT     T1528 K20
      AND     T1528
      SET     M1782
      RST     M1792
      AND>    D1655 K0
      DEC     D1655
15    LD      M1791
      SET     M1750
      SET     M1792
      RST     M1791
19    LD      M1790
      ANI     M1750
      AND     M1886
      LDI     M1751
      ORI     M1800
      ANB
      SET     M1791
      RST     M1790
      AND     M1751
      SET     M1754
29    LD      M1789
      SET     M1953
      SET     M1752
      SET     M1788
      RST     M1789
34    LD      M1788
      SET     M1790
      RST     M1788
      LD      M1752
      OR<>    D1700 K1
      ANB
      SET     M1751
43    LD      M1787
      SET     M1953
      SET     M1786
      RST     M1787
47    LD      M1786
      MOV     K0 D1710
      SET     M1788
      RST     M1786
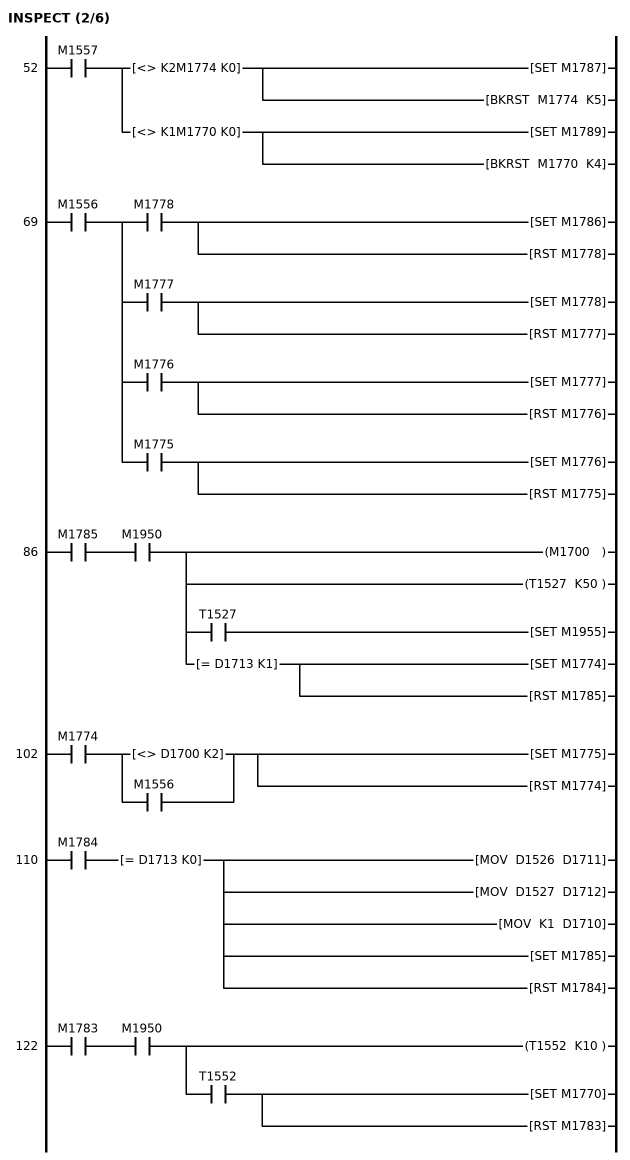
52    LD      M1557
      MPS
      AND<>   K2M1774 K0
      SET     M1787
      BKRST   M1774 K5
      MPP
      AND<>   K1M1770 K0
      SET     M1789
      BKRST   M1770 K4
69    LD      M1556
      MPS
      AND     M1778
      SET     M1786
      RST     M1778
      MRD
      AND     M1777
      SET     M1778
      RST     M1777
      MRD
      AND     M1776
      SET     M1777
      RST     M1776
      MPP
      AND     M1775
      SET     M1776
      RST     M1775
86    LD      M1785
      AND     M1950
      OUT     M1700
      OUT     T1527 K50
      MPS
      AND     T1527
      SET     M1955
      MPP
      AND=    D1713 K1
      SET     M1774
      RST     M1785
102   LD      M1774
      LD<>    D1700 K2
      OR      M1556
      ANB
      SET     M1775
      RST     M1774
110   LD      M1784
      AND=    D1713 K0
      MOV     D1526 D1711
      MOV     D1527 D1712
      MOV     K1 D1710
      SET     M1785
      RST     M1784
122   LD      M1783
      AND     M1950
      OUT     T1552 K10
      AND     T1552
      SET     M1770
      RST     M1783
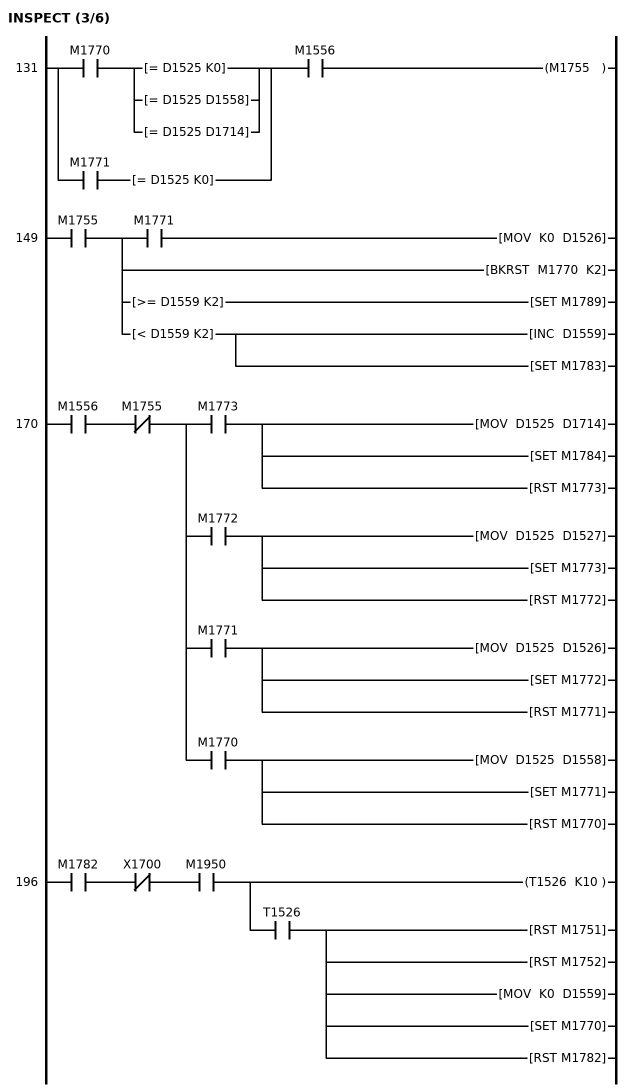
131   LD      M1770
      LD=     D1525 K0
      OR=     D1525 D1558
      OR=     D1525 D1714
      ANB
      LD      M1771
      AND=    D1525 K0
      ORB
      AND     M1556
      OUT     M1755
149   LD      M1755
      MPS
      AND     M1771
      MOV     K0 D1526
      MPP
      BKRST   M1770 K2
      MPS
      AND>=   D1559 K2
      SET     M1789
      MPP
      AND<    D1559 K2
      INC     D1559
      SET     M1783
170   LD      M1556
      ANI     M1755
      MPS
      AND     M1773
      MOV     D1525 D1714
      SET     M1784
      RST     M1773
      MRD
      AND     M1772
      MOV     D1525 D1527
      SET     M1773
      RST     M1772
      MRD
      AND     M1771
      MOV     D1525 D1526
      SET     M1772
      RST     M1771
      MPP
      AND     M1770
      MOV     D1525 D1558
      SET     M1771
      RST     M1770
196   LD      M1782
      ANI     X1700
      AND     M1950
      OUT     T1526 K10
      AND     T1526
      RST     M1751
      RST     M1752
      MOV     K0 D1559
      SET     M1770
      RST     M1782
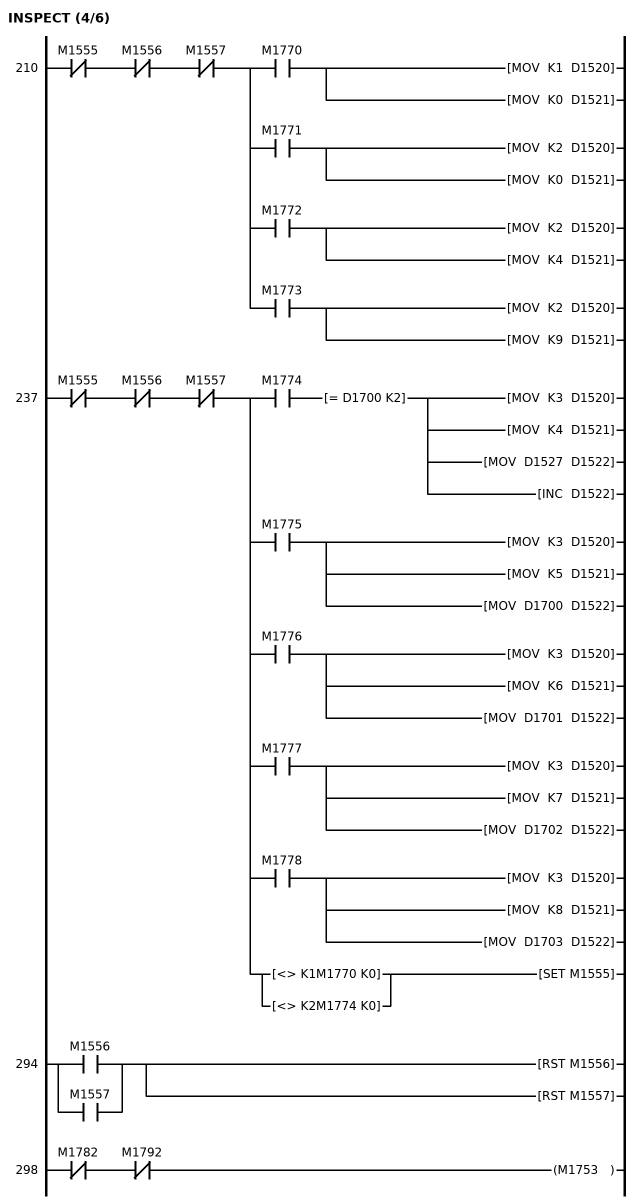
210   LDI     M1555
      ANI     M1556
      ANI     M1557
      MPS
      AND     M1770
      MOV     K1 D1520
      MOV     K0 D1521
      MRD
      AND     M1771
      MOV     K2 D1520
      MOV     K0 D1521
      MRD
      AND     M1772
      MOV     K2 D1520
      MOV     K4 D1521
      MPP
      AND     M1773
      MOV     K2 D1520
      MOV     K9 D1521
237   LDI     M1555
      ANI     M1556
      ANI     M1557
      MPS
      AND     M1774
      AND=    D1700 K2
      MOV     K3 D1520
      MOV     K4 D1521
      MOV     D1527 D1522
      INC     D1522
      MRD
      AND     M1775
      MOV     K3 D1520
      MOV     K5 D1521
      MOV     D1700 D1522
      MRD
      AND     M1776
      MOV     K3 D1520
      MOV     K6 D1521
      MOV     D1701 D1522
      MRD
      AND     M1777
      MOV     K3 D1520
      MOV     K7 D1521
      MOV     D1702 D1522
      MRD
      AND     M1778
      MOV     K3 D1520
      MOV     K8 D1521
      MOV     D1703 D1522
      MPP
      LD<>    K1M1770 K0
      OR<>    K2M1774 K0
      ANB
      SET     M1555
294   LD      M1556
      OR      M1557
      RST     M1556
      RST     M1557
298   LDI     M1782
      ANI     M1792
      OUT     M1753
